(* IEC 61131-3 sources: Gen-AI/final/Gen-AI_v1.0_submission/A2_框架源码/agent/logs/scenario_fixture/best-effort/fixture/E3_S02_1_42, 3 files *)

(* ---- best.st ---- *)
FUNCTION_BLOCK FB_S02
VAR_INPUT
    FwdBtn : BOOL;
    RevBtn : BOOL;
    MaintKey : BOOL;
    EStop_NC : BOOL;
END_VAR
VAR_OUTPUT
    MotorFwd : BOOL;
    MotorRev : BOOL;
    RunLamp : BOOL;
    Status : WORD;
END_VAR
(* Add a VAR block for internal state/timers before the implementation, if needed. *)
(* SKELETON ONLY: replace this RETURN with scan logic and required initial state. *)
RETURN;
END_FUNCTION_BLOCK

(* FIXTURE_TEST_FAIL *)

(* ---- final.st ---- *)
FUNCTION_BLOCK FB_S02
VAR_INPUT
    FwdBtn : BOOL;
    RevBtn : BOOL;
    MaintKey : BOOL;
    EStop_NC : BOOL;
END_VAR
VAR_OUTPUT
    MotorFwd : BOOL;
    MotorRev : BOOL;
    RunLamp : BOOL;
    Status : WORD;
END_VAR
(* Add a VAR block for internal state/timers before the implementation, if needed. *)
(* SKELETON ONLY: replace this RETURN with scan logic and required initial state. *)
RETURN;
END_FUNCTION_BLOCK

(* FIXTURE_TEST_FAIL *)

(* ---- skeleton.st ---- *)
FUNCTION_BLOCK FB_S02
VAR_INPUT
    FwdBtn : BOOL;
    RevBtn : BOOL;
    MaintKey : BOOL;
    EStop_NC : BOOL;
END_VAR
VAR_OUTPUT
    MotorFwd : BOOL;
    MotorRev : BOOL;
    RunLamp : BOOL;
    Status : WORD;
END_VAR
(* Add a VAR block for internal state/timers before the implementation, if needed. *)
(* SKELETON ONLY: replace this RETURN with scan logic and required initial state. *)
RETURN;
END_FUNCTION_BLOCK
